(*
SPDX-FileCopyrightText: c 2026 Oleksandr Tiutyk <trofimich@gmail.com>
SPDX-License-Identifier: MIT
License: https://opensource.org/license/mit
*)

(*!
<summary>Groups fixed-capacity stack storage, LIFO order, cursors, ownership and overflow cases.</summary>
<description>
Owns the cases, their fixed registration array and any fixtures borrowed by the cases.
Each borrowed fixture is reserved for its case throughout the group lifetime. Use from one task at a stable address.
</description>
*)

{attribute 'no_assign'}
{attribute 'no_explicit_call' := 'do not call this function block directly'}
FUNCTION_BLOCK StaticStackTestGroup EXTENDS TOF_Testing.TestGroup<11>
VAR_STAT
	{attribute 'hide'}
	_ClassName : STRING := __POUNAME();
END_VAR
VAR
	_Validator : TOF_Core.GenericValueTypeValidator(typeClass := TOF_Core.GENERIC_TYPE_CLASS.INT_16);
	_OwnedObjectCleanupStack : TOF_Collections.Stack<3>(valueValidator := 0);
	_ValidatorRejectionStack : TOF_Collections.Stack<3>(valueValidator := _Validator);
	_IndexedAccessAndEnumerationStack : TOF_Collections.Stack<3>(valueValidator := 0);
	_EmptyAndIndexBoundsStack : TOF_Collections.Stack<3>(valueValidator := 0);
	_CopiedAndBorrowedValuesStack : TOF_Collections.Stack<3>(valueValidator := 0);
	_ContainsStack : TOF_Collections.Stack<3>(valueValidator := 0);
	_ContainsGenericStack : TOF_Collections.Stack<3>(valueValidator := 0);
	_PushAndPeekStack : TOF_Collections.Stack<3>(valueValidator := 0);
	_RemoveLastStack : TOF_Collections.Stack<3>(valueValidator := 0);

	_OwnedObjectCleanup : StackOwnedObjectCleanupTest(
		name := "OwnedObjectCleanup",
		parent := THIS^,
		stack := _OwnedObjectCleanupStack
	);
	_ValidatorRejection : StackValidatorRejectionTest(
		name := "ValidatorRejection",
		parent := THIS^,
		stack := _ValidatorRejectionStack
	);
	_IndexedAccessAndEnumeration : StackIndexedAccessAndEnumerationTest(
		name := "IndexedAccessAndEnumeration",
		parent := THIS^,
		stack := _IndexedAccessAndEnumerationStack
	);
	_EmptyAndIndexBounds : StackEmptyAndIndexBoundsTest(
		name := "EmptyAndIndexBounds",
		parent := THIS^,
		stack := _EmptyAndIndexBoundsStack
	);
	_CopiedAndBorrowedValues : StackCopiedAndBorrowedValuesTest(
		name := "CopiedAndBorrowedValues",
		parent := THIS^,
		stack := _CopiedAndBorrowedValuesStack
	);
	_Contains : StackContainsTest(name := "Contains", parent := THIS^, stack := _ContainsStack);
	_ContainsGeneric : StackContainsGenericTest(
		name := "ContainsGeneric",
		parent := THIS^,
		stack := _ContainsGenericStack
	);
	_PushAndPeek : StackPushAndPeekTest(name := "PushAndPeek", parent := THIS^, stack := _PushAndPeekStack);
	_Clear : StaticStackClearTest(name := "Clear", parent := THIS^);
	_RemoveLast : StackRemoveLastTest(name := "RemoveLast", parent := THIS^, stack := _RemoveLastStack);
	_Overflow : StaticStackOverflowTest(name := "Overflow", parent := THIS^);

	_Children : ARRAY [0.._ChildCount - 1] OF TOF_Testing.ITestElement :=
	[
		_OwnedObjectCleanup,
		_ValidatorRejection,
		_IndexedAccessAndEnumeration,
		_EmptyAndIndexBounds,
		_CopiedAndBorrowedValues,
		_Contains,
		_ContainsGeneric,
		_PushAndPeek,
		_Clear,
		_RemoveLast,
		_Overflow
	];
END_VAR

//! <summary>Borrows the fixed child array. Callers must not modify it.</summary>
{attribute 'monitoring' := 'call'}
PROPERTY Children : REFERENCE TO ARRAY [0.._ChildCount - 1] OF TOF_Testing.ITestElement
GET
Children REF= _Children;
END_GET
END_PROPERTY

//! <summary>Borrows the concrete class name. Callers must not modify it.</summary>
{attribute 'monitoring' := 'call'}
PROPERTY ClassName : REFERENCE TO STRING
GET
ClassName REF= _ClassName;
END_GET
END_PROPERTY

//! <summary>Borrows the compiler-initialized namespace name. Callers must not modify it.</summary>
{attribute 'monitoring' := 'call'}
PROPERTY NamespaceName : REFERENCE TO STRING
GET
NamespaceName REF= CurrentNamespace.Name;
END_GET
END_PROPERTY

//! <summary>Reports the concrete instance size in bytes.</summary>
{attribute 'monitoring' := 'call'}
PROPERTY SelfSize : ULINT
GET
SelfSize := XSIZEOF(THIS^);
END_GET
END_PROPERTY

END_FUNCTION_BLOCK

(* stored: Version 1.1.0.1
   POU StaticStackTestGroup: Id {8848843b-576f-4850-8977-11e8bc08bd08}, SpecialFunc None
   Property Children: Id {16e7fb71-bd9e-4fa6-b41a-3fb4546cb480}
   Get Get: Id {fe862984-5a29-4389-af09-a7cc710be9e0}
   Property ClassName: Id {0414519b-5039-4831-94f1-efee7df3b69f}
   Get Get: Id {571e0a77-546b-4707-9912-878c2f82e2ac}
   Property NamespaceName: Id {119d2abd-e05a-4abf-9fd4-d773ab40c1c0}
   Get Get: Id {22ed5e41-5655-46ed-a4ce-2f78b9e79255}
   Property SelfSize: Id {65649c38-40c4-4d8b-b867-34d139c4d035}
   Get Get: Id {3cc5b5da-ee02-4a72-9772-3d1723144d6e} *)
